Fanuc KAREL source: ks00040.KL

PROGRAM KS00040
%STACKSIZE=65535
%PRIORITY=65535
%NOLOCKGROUP
VAR
A : ARRAY[4] OF POSITION
B : ARRAY[4] OF POSITION
FLAG : BOOLEAN
N : INTEGER
STATUS : INTEGER
PN : STRING[80]
VN : STRING[80]
BEGIN
PN=''
VN='A'
-- UNSAFE_SOURCE_IR line 19: N = native_s16_value(A)
END KS00040
